Staubli VAL3: create.pgx

public program create()
begin
  call init()
  //action control management
  taskKill("actCtrl")
  taskCreate "actCtrl",100,_tActCtrl()
  wait(taskStatus("actCtrl")==1)
end
